(* IEC 61131-3 sources: llm-plc-st-eval/data/processed_v2_primera/gpt-4o/I4/few_shot, 3 files *)

(* ---- ejec_1.st ---- *)
FUNCTION_BLOCK FB_EstrellaTriangulo
VAR_INPUT
    btnMarcha : BOOL; (* Botón de marcha *)
    btnParo : BOOL;   (* Botón de paro *)
END_VAR
VAR_OUTPUT
    kM : BOOL; (* Contactor principal *)
    kY : BOOL; (* Contactor de estrella *)
    kD : BOOL; (* Contactor de triángulo *)
END_VAR
VAR
    tEstrella : TON; (* Temporizador para estrella *)
    tTiempoMuerto : TON; (* Temporizador para tiempo muerto *)
    estado : INT; (* Estado del arranque *)
END_VAR

(* Lógica de control de arranque estrella-triángulo *)
IF btnParo THEN
    (* Reset de todos los contactores y temporizadores en caso de paro *)
    kM := FALSE;
    kY := FALSE;
    kD := FALSE;
    tEstrella(IN := FALSE);
    tTiempoMuerto(IN := FALSE);
    estado := 0;
ELSIF btnMarcha THEN
    CASE estado OF
        0: (* Estado inicial, activa contactor principal y estrella *)
            kM := TRUE;
            kY := TRUE;
            tEstrella(IN := TRUE, PT := T#8S);
            estado := 1;
        1: (* Espera el tiempo de estrella *)
            IF tEstrella.Q THEN
                kY := FALSE;
                tTiempoMuerto(IN := TRUE, PT := T#100MS);
                estado := 2;
            END_IF
        2: (* Espera el tiempo muerto *)
            IF tTiempoMuerto.Q THEN
                kD := TRUE;
                estado := 3;
            END_IF
        3: (* Estado final, solo contactor de triángulo activo *)
            (* Mantener kM y kD activos *)
    END_CASE
ELSE
    (* Si no hay marcha ni paro, desactivar todos los contactores *)
    kM := FALSE;
    kY := FALSE;
    kD := FALSE;
    tEstrella(IN := FALSE);
    tTiempoMuerto(IN := FALSE);
    estado := 0;
END_IF
END_FUNCTION_BLOCK

(* ---- ejec_2.st ---- *)
FUNCTION_BLOCK FB_EstrellaTriangulo
VAR_INPUT
    btnMarcha : BOOL; (* Botón de marcha *)
    btnParo : BOOL;   (* Botón de paro *)
END_VAR
VAR_OUTPUT
    kM : BOOL; (* Contactor principal *)
    kY : BOOL; (* Contactor de estrella *)
    kD : BOOL; (* Contactor de triángulo *)
END_VAR
VAR
    timerEstrella : TON; (* Temporizador para estrella *)
    timerMuerto : TON;   (* Temporizador para tiempo muerto *)
    estado : INT;        (* Estado del arranque *)
END_VAR

(* Lógica de control del arranque estrella-triángulo *)
IF btnParo THEN
    (* Reset de todos los contactores y temporizadores al pulsar paro *)
    kM := FALSE;
    kY := FALSE;
    kD := FALSE;
    timerEstrella(IN := FALSE);
    timerMuerto(IN := FALSE);
    estado := 0;
ELSIF btnMarcha THEN
    CASE estado OF
        0: (* Estado inicial, activa contactor principal y estrella *)
            kM := TRUE;
            kY := TRUE;
            timerEstrella(IN := TRUE, PT := T#8S);
            estado := 1;
        1: (* Espera tiempo de estrella *)
            IF timerEstrella.Q THEN
                kY := FALSE;
                timerMuerto(IN := TRUE, PT := T#100MS);
                estado := 2;
            END_IF
        2: (* Espera tiempo muerto *)
            IF timerMuerto.Q THEN
                kD := TRUE;
                estado := 3;
            END_IF
        3: (* Estado final, contactor de triángulo activado *)
            (* Mantener kM y kD activados *)
    END_CASE
ELSE
    (* Si no se pulsa marcha, reset de todos los contactores y temporizadores *)
    kM := FALSE;
    kY := FALSE;
    kD := FALSE;
    timerEstrella(IN := FALSE);
    timerMuerto(IN := FALSE);
    estado := 0;
END_IF
END_FUNCTION_BLOCK

(* ---- ejec_3.st ---- *)
FUNCTION_BLOCK FB_EstrellaTriangulo
VAR_INPUT
    btnMarcha : BOOL; (* Botón de marcha *)
    btnParo : BOOL;   (* Botón de paro *)
END_VAR
VAR_OUTPUT
    kM : BOOL; (* Contactor principal *)
    kY : BOOL; (* Contactor estrella *)
    kD : BOOL; (* Contactor triángulo *)
END_VAR
VAR
    tEstrella : TON;  (* Temporizador para estrella *)
    tMuerto : TON;    (* Temporizador para tiempo muerto *)
    estado : INT;     (* Estado del arranque *)
END_VAR

(* Lógica de control del arranque estrella-triángulo *)
IF btnParo THEN
    (* Si se presiona el botón de paro, desactivar todos los contactores *)
    kM := FALSE;
    kY := FALSE;
    kD := FALSE;
    estado := 0;
ELSIF btnMarcha THEN
    CASE estado OF
        0: (* Estado inicial, activar contactor principal y estrella *)
            kM := TRUE;
            kY := TRUE;
            tEstrella(IN := TRUE, PT := T#8S);
            estado := 1;
        1: (* Esperar 8 segundos con contactor estrella activado *)
            IF tEstrella.Q THEN
                kY := FALSE; (* Desactivar contactor estrella *)
                tMuerto(IN := TRUE, PT := T#100MS);
                estado := 2;
            END_IF
        2: (* Esperar tiempo muerto de 100 ms *)
            IF tMuerto.Q THEN
                kD := TRUE; (* Activar contactor triángulo *)
                estado := 3;
            END_IF
        3: (* Estado final, contactor triángulo activado *)
            (* Mantener estado hasta que se presione btnParo *)
    END_CASE
ELSE
    (* Si no se presiona ningún botón, mantener estado actual *)
    tEstrella(IN := FALSE);
    tMuerto(IN := FALSE);
END_IF
END_FUNCTION_BLOCK
